KUKA KRL program: ManyMoves.src

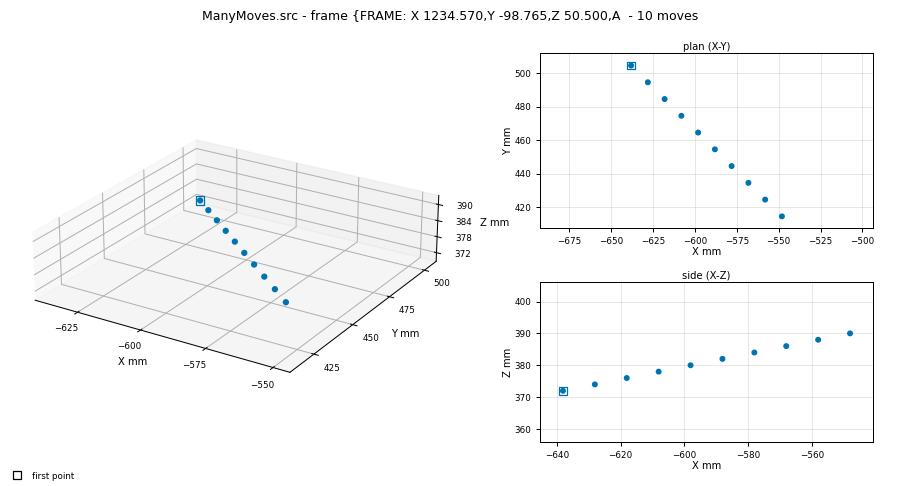
[picture p0: tool path of ManyMoves.src in frame {FRAME: X 1234.570,Y -98.765,Z 50.500,A , 10 of 30 moves have a stored position in this frame; points joined in program order, loops and branches not executed]
&ACCESS RVP
&REL 1
&PARAM TEMPLATE = C:\KRC\Roboter\Template\vorgabe
&PARAM EDITMASK = *
DEF ManyMoves ( )


; GLOBAL INTERRUPT DECL 3 WHEN $STOPMESS==TRUE DO IR_STOPM ( )
; INTERRUPT ON 3

;FOLD Initialise and set default speed
BAS (#INITMOV,0)
BAS (#VEL_PTP,100)
BAS (#ACC_PTP,20)
$VEL.CP=0.2
BAS (#TOOL,0)
BAS (#BASE,0)
;ENDFOLD

;;FOLD STARTPOS
;$BWDSTART = FALSE
;PDAT_ACT = PDEFAULT
;BAS(#PTP_DAT)
;FDAT_ACT = {TOOL_NO 0,BASE_NO 0,IPO_FRAME #BASE}
;BAS(#FRAMES)
;;ENDFOLD

$ADVANCE = 5

;FOLD ---- Quickly skip BCO ----
; PTP $AXIS_ACT
;ENDFOLD

;FOLD ---- GO HOME ----
; PTP {A1 0.000, A2 -90.000, A3 90.000, A4 0.000, A5 0.000, A6 0.000, E1 0, E2 0, E3 0, E4 0, E5 0, E6 0}
;ENDFOLD


; Program generated by RoboDK v6.0.7 for KUKA IONTEC ultra KR 120 R2700 on XX/XX/XXXX 18:00:00
; Using nominal kinematics.
; ---- Setting reference (Base) ----
$BASE = {FRAME: X 1234.570,Y -98.765,Z 50.500,A 30.000,B 0.000,C 0.000}
; --------------------------
; ---- Setting tool (TCP) ----
$TOOL = {FRAME: X 10.000,Y 20.000,Z 150.000,A 0.000,B 0.000,C 0.000}
; --------------------------
$VEL.CP = 0.50000
PTP {A1 0.00000,A2 -10.00000,A3 20.00000,A4 0.00000,A5 30.00000,A6 0.00000}
LIN {X -638.084,Y 504.480,Z 372.034,A 150.000,B 50.000,C -165.000}
PTP {A1 20.00000,A2 -10.00000,A3 20.00000,A4 0.00000,A5 30.00000,A6 0.00000}
; Linear movement using joint targets is not supported. Change the target type to cartesian or use a joint movement.
PTP {A1 0.00000,A2 -10.00000,A3 20.00000,A4 0.00000,A5 30.00000,A6 0.00000}
LIN {X -628.084,Y 494.480,Z 374.034,A 150.000,B 50.000,C -165.000}
PTP {A1 20.00000,A2 -10.00000,A3 20.00000,A4 0.00000,A5 30.00000,A6 0.00000}
; Linear movement using joint targets is not supported. Change the target type to cartesian or use a joint movement.
PTP {A1 0.00000,A2 -10.00000,A3 20.00000,A4 0.00000,A5 30.00000,A6 0.00000}
LIN {X -618.084,Y 484.480,Z 376.034,A 150.000,B 50.000,C -165.000}
PTP {A1 20.00000,A2 -10.00000,A3 20.00000,A4 0.00000,A5 30.00000,A6 0.00000}
; Linear movement using joint targets is not supported. Change the target type to cartesian or use a joint movement.
PTP {A1 0.00000,A2 -10.00000,A3 20.00000,A4 0.00000,A5 30.00000,A6 0.00000}
LIN {X -608.084,Y 474.480,Z 378.034,A 150.000,B 50.000,C -165.000}
PTP {A1 20.00000,A2 -10.00000,A3 20.00000,A4 0.00000,A5 30.00000,A6 0.00000}
; Linear movement using joint targets is not supported. Change the target type to cartesian or use a joint movement.
PTP {A1 0.00000,A2 -10.00000,A3 20.00000,A4 0.00000,A5 30.00000,A6 0.00000}
LIN {X -598.084,Y 464.480,Z 380.034,A 150.000,B 50.000,C -165.000}
PTP {A1 20.00000,A2 -10.00000,A3 20.00000,A4 0.00000,A5 30.00000,A6 0.00000}
; Linear movement using joint targets is not supported. Change the target type to cartesian or use a joint movement.
PTP {A1 0.00000,A2 -10.00000,A3 20.00000,A4 0.00000,A5 30.00000,A6 0.00000}
LIN {X -588.084,Y 454.480,Z 382.034,A 150.000,B 50.000,C -165.000}
PTP {A1 20.00000,A2 -10.00000,A3 20.00000,A4 0.00000,A5 30.00000,A6 0.00000}
; Linear movement using joint targets is not supported. Change the target type to cartesian or use a joint movement.
PTP {A1 0.00000,A2 -10.00000,A3 20.00000,A4 0.00000,A5 30.00000,A6 0.00000}
LIN {X -578.084,Y 444.480,Z 384.034,A 150.000,B 50.000,C -165.000}
PTP {A1 20.00000,A2 -10.00000,A3 20.00000,A4 0.00000,A5 30.00000,A6 0.00000}
; Linear movement using joint targets is not supported. Change the target type to cartesian or use a joint movement.
PTP {A1 0.00000,A2 -10.00000,A3 20.00000,A4 0.00000,A5 30.00000,A6 0.00000}
LIN {X -568.084,Y 434.480,Z 386.034,A 150.000,B 50.000,C -165.000}
PTP {A1 20.00000,A2 -10.00000,A3 20.00000,A4 0.00000,A5 30.00000,A6 0.00000}
; Linear movement using joint targets is not supported. Change the target type to cartesian or use a joint movement.
PTP {A1 0.00000,A2 -10.00000,A3 20.00000,A4 0.00000,A5 30.00000,A6 0.00000}
LIN {X -558.084,Y 424.480,Z 388.034,A 150.000,B 50.000,C -165.000}
PTP {A1 20.00000,A2 -10.00000,A3 20.00000,A4 0.00000,A5 30.00000,A6 0.00000}
; Linear movement using joint targets is not supported. Change the target type to cartesian or use a joint movement.
PTP {A1 0.00000,A2 -10.00000,A3 20.00000,A4 0.00000,A5 30.00000,A6 0.00000}
LIN {X -548.084,Y 414.480,Z 390.034,A 150.000,B 50.000,C -165.000}
PTP {A1 20.00000,A2 -10.00000,A3 20.00000,A4 0.00000,A5 30.00000,A6 0.00000}
; Linear movement using joint targets is not supported. Change the target type to cartesian or use a joint movement.
END
